Fanuc KAREL source: kc00005.KL

-- PROVISIONAL review KL for V770-1; original PC SHA256 8509346717ef151aeb61727a2e23bdc0729c98ecce21cdb6a2b3436b8e75ced9
-- Incomplete behavior may be omitted. Consult companion uncertainty JSON. Do not deploy.
PROGRAM KC00005
%NOLOCKGROUP
BEGIN
  -- UNRESOLVED_PC offsets 5-27; opcodes 27,22,22,22,31
  -- UNRESOLVED_PC offsets 32-36; opcodes 7F
END KC00005
